Staubli VAL3: setDigOutput.pgx

public program setDigOutput(dio& x_dOut, bool x_bValue, bool& x_bError)
  local string l_sDesc
  local string l_sPath
begin
  if ioStatus(x_dOut,l_sDesc,l_sPath)>=0
    x_bError=false
    x_dOut=x_bValue
  else
    x_bError=true
//    logMsg("Signal "+l_sPath+" error."+"Description:"+l_sDesc)
  endIf

end
